// Who may command the telescope: the physical Local/Remote switch (or the fixed project policy). I_Cabinet.ControlMode.
{attribute 'qualified_only'}
{attribute 'strict'}
TYPE E_ControlMode :
(
	remote := 0,
	local := 1
);
END_TYPE

(* stored: Version 1.1.0.1, ProductVersion 3.1.4024.15
   DUT E_ControlMode: Id {21390704-2bb3-46ec-bebb-9447898de08a} *)
